Universal Robots URScript: horizontal_swab_path.script

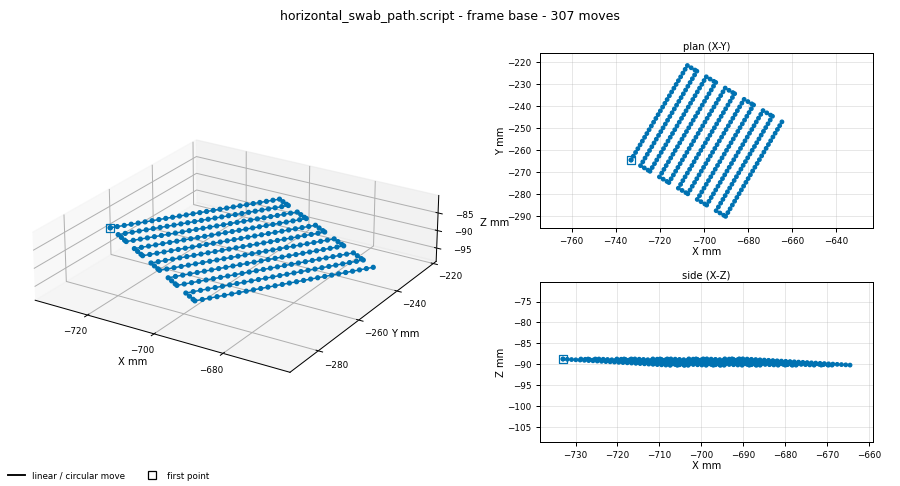
[picture p0: tool path of horizontal_swab_path.script in frame base, 307 of 307 moves have a stored position in this frame; points joined in program order, loops and branches not executed]
def horizontal_swab_path():

  # Move to first swab point perpendicular
  movel(p[-0.73300831, -0.26450111, -0.08872548, -0.83237244, -3.02179964, 0.04578505], a=0.2000, v=0.0300, r=0.0000)

  # Incline tool while keeping TCP XYZ fixed
  movel(p[-0.73300831, -0.26450111, -0.08872548, -0.64311438, -2.27932698, -0.22586576], a=0.1000, v=0.0150, r=0.0000)
  # Horizontal waypoint 1
  movel(p[-0.73198462, -0.26278399, -0.08878548, -0.64311438, -2.27932698, -0.22586576], a=0.1500, v=0.0200, r=0.0000)
  # Horizontal waypoint 2
  movel(p[-0.73096094, -0.26106688, -0.08884547, -0.64311438, -2.27932698, -0.22586576], a=0.1500, v=0.0200, r=0.0000)
  # Horizontal waypoint 3
  movel(p[-0.72993725, -0.25934977, -0.08890546, -0.64311438, -2.27932698, -0.22586576], a=0.1500, v=0.0200, r=0.0000)
  # Horizontal waypoint 4
  movel(p[-0.72891357, -0.25763266, -0.08896545, -0.64311438, -2.27932698, -0.22586576], a=0.1500, v=0.0200, r=0.0000)
  # Horizontal waypoint 5
  movel(p[-0.72788988, -0.25591555, -0.08902544, -0.64311438, -2.27932698, -0.22586576], a=0.1500, v=0.0200, r=0.0000)
  # Horizontal waypoint 6
  movel(p[-0.72686620, -0.25419844, -0.08908543, -0.64311438, -2.27932698, -0.22586576], a=0.1500, v=0.0200, r=0.0000)
  # Horizontal waypoint 7
  movel(p[-0.72584251, -0.25248133, -0.08914542, -0.64311438, -2.27932698, -0.22586576], a=0.1500, v=0.0200, r=0.0000)
  # Horizontal waypoint 8
  movel(p[-0.72481883, -0.25076422, -0.08920541, -0.64311438, -2.27932698, -0.22586576], a=0.1500, v=0.0200, r=0.0000)
  # Horizontal waypoint 9
  movel(p[-0.72379514, -0.24904710, -0.08926540, -0.64311438, -2.27932698, -0.22586576], a=0.1500, v=0.0200, r=0.0000)
  # Horizontal waypoint 10
  movel(p[-0.72277146, -0.24732999, -0.08932539, -0.64311438, -2.27932698, -0.22586576], a=0.1500, v=0.0200, r=0.0000)
  # Horizontal waypoint 11
  movel(p[-0.72174777, -0.24561288, -0.08938538, -0.64311438, -2.27932698, -0.22586576], a=0.1500, v=0.0200, r=0.0000)
  # Horizontal waypoint 12
  movel(p[-0.72072409, -0.24389577, -0.08944538, -0.64311438, -2.27932698, -0.22586576], a=0.1500, v=0.0200, r=0.0000)
  # Horizontal waypoint 13
  movel(p[-0.71970040, -0.24217866, -0.08950537, -0.64311438, -2.27932698, -0.22586576], a=0.1500, v=0.0200, r=0.0000)
  # Horizontal waypoint 14
  movel(p[-0.71867672, -0.24046155, -0.08956536, -0.64311438, -2.27932698, -0.22586576], a=0.1500, v=0.0200, r=0.0000)
  # Horizontal waypoint 15
  movel(p[-0.71765303, -0.23874444, -0.08962535, -0.64311438, -2.27932698, -0.22586576], a=0.1500, v=0.0200, r=0.0000)
  # Horizontal waypoint 16
  movel(p[-0.71662935, -0.23702733, -0.08968534, -0.64311438, -2.27932698, -0.22586576], a=0.1500, v=0.0200, r=0.0000)
  # Horizontal waypoint 17
  movel(p[-0.71560566, -0.23531022, -0.08974533, -0.64311438, -2.27932698, -0.22586576], a=0.1500, v=0.0200, r=0.0000)
  # Horizontal waypoint 18
  movel(p[-0.71458198, -0.23359311, -0.08980532, -0.64311438, -2.27932698, -0.22586576], a=0.1500, v=0.0200, r=0.0000)
  # Horizontal waypoint 19
  movel(p[-0.71355829, -0.23187600, -0.08986531, -0.64311438, -2.27932698, -0.22586576], a=0.1500, v=0.0200, r=0.0000)
  # Horizontal waypoint 20
  movel(p[-0.71253461, -0.23015888, -0.08992530, -0.64311438, -2.27932698, -0.22586576], a=0.1500, v=0.0200, r=0.0000)
  # Horizontal waypoint 21
  movel(p[-0.71151092, -0.22844177, -0.08998530, -0.64311438, -2.27932698, -0.22586576], a=0.1500, v=0.0200, r=0.0000)
  # Horizontal waypoint 22
  movel(p[-0.71048724, -0.22672466, -0.09004529, -0.64311438, -2.27932698, -0.22586576], a=0.1500, v=0.0200, r=0.0000)
  # Horizontal waypoint 23
  movel(p[-0.70946356, -0.22500755, -0.09010528, -0.64311438, -2.27932698, -0.22586576], a=0.1500, v=0.0200, r=0.0000)
  # Horizontal waypoint 24
  movel(p[-0.70843987, -0.22329044, -0.09016527, -0.64311438, -2.27932698, -0.22586576], a=0.1500, v=0.0200, r=0.0000)
  # Horizontal waypoint 25
  movel(p[-0.70741619, -0.22157333, -0.09022526, -0.64311438, -2.27932698, -0.22586576], a=0.1500, v=0.0200, r=0.0000)
  # Horizontal waypoint 26
  movel(p[-0.70569827, -0.22259742, -0.09022307, -0.64311438, -2.27932698, -0.22586576], a=0.1500, v=0.0200, r=0.0000)
  # Horizontal waypoint 27
  movel(p[-0.70398035, -0.22362151, -0.09022089, -0.64311438, -2.27932698, -0.22586576], a=0.1500, v=0.0200, r=0.0000)
  # Horizontal waypoint 28
  movel(p[-0.70312139, -0.22413355, -0.09021980, -0.64311438, -2.27932698, -0.22586576], a=0.1500, v=0.0200, r=0.0000)
  # Horizontal waypoint 29
  movel(p[-0.70414508, -0.22585066, -0.09015981, -0.64311438, -2.27932698, -0.22586576], a=0.1500, v=0.0200, r=0.0000)
  # Horizontal waypoint 30
  movel(p[-0.70516876, -0.22756777, -0.09009982, -0.64311438, -2.27932698, -0.22586576], a=0.1500, v=0.0200, r=0.0000)
  # Horizontal waypoint 31
  movel(p[-0.70619245, -0.22928488, -0.09003983, -0.64311438, -2.27932698, -0.22586576], a=0.1500, v=0.0200, r=0.0000)
  # Horizontal waypoint 32
  movel(p[-0.70721613, -0.23100199, -0.08997983, -0.64311438, -2.27932698, -0.22586576], a=0.1500, v=0.0200, r=0.0000)
  # Horizontal waypoint 33
  movel(p[-0.70823982, -0.23271911, -0.08991984, -0.64311438, -2.27932698, -0.22586576], a=0.1500, v=0.0200, r=0.0000)
  # Horizontal waypoint 34
  movel(p[-0.70926350, -0.23443622, -0.08985985, -0.64311438, -2.27932698, -0.22586576], a=0.1500, v=0.0200, r=0.0000)
  # Horizontal waypoint 35
  movel(p[-0.71028719, -0.23615333, -0.08979986, -0.64311438, -2.27932698, -0.22586576], a=0.1500, v=0.0200, r=0.0000)
  # Horizontal waypoint 36
  movel(p[-0.71131087, -0.23787044, -0.08973987, -0.64311438, -2.27932698, -0.22586576], a=0.1500, v=0.0200, r=0.0000)
  # Horizontal waypoint 37
  movel(p[-0.71233456, -0.23958755, -0.08967988, -0.64311438, -2.27932698, -0.22586576], a=0.1500, v=0.0200, r=0.0000)
  # Horizontal waypoint 38
  movel(p[-0.71335824, -0.24130466, -0.08961989, -0.64311438, -2.27932698, -0.22586576], a=0.1500, v=0.0200, r=0.0000)
  # Horizontal waypoint 39
  movel(p[-0.71438193, -0.24302177, -0.08955990, -0.64311438, -2.27932698, -0.22586576], a=0.1500, v=0.0200, r=0.0000)
  # Horizontal waypoint 40
  movel(p[-0.71540561, -0.24473888, -0.08949991, -0.64311438, -2.27932698, -0.22586576], a=0.1500, v=0.0200, r=0.0000)
  # Horizontal waypoint 41
  movel(p[-0.71642930, -0.24645599, -0.08943991, -0.64311438, -2.27932698, -0.22586576], a=0.1500, v=0.0200, r=0.0000)
  # Horizontal waypoint 42
  movel(p[-0.71745298, -0.24817311, -0.08937992, -0.64311438, -2.27932698, -0.22586576], a=0.1500, v=0.0200, r=0.0000)
  # Horizontal waypoint 43
  movel(p[-0.71847667, -0.24989022, -0.08931993, -0.64311438, -2.27932698, -0.22586576], a=0.1500, v=0.0200, r=0.0000)
  # Horizontal waypoint 44
  movel(p[-0.71950035, -0.25160733, -0.08925994, -0.64311438, -2.27932698, -0.22586576], a=0.1500, v=0.0200, r=0.0000)
  # Horizontal waypoint 45
  movel(p[-0.72052404, -0.25332444, -0.08919995, -0.64311438, -2.27932698, -0.22586576], a=0.1500, v=0.0200, r=0.0000)
  # Horizontal waypoint 46
  movel(p[-0.72154772, -0.25504155, -0.08913996, -0.64311438, -2.27932698, -0.22586576], a=0.1500, v=0.0200, r=0.0000)
  # Horizontal waypoint 47
  movel(p[-0.72257141, -0.25675866, -0.08907997, -0.64311438, -2.27932698, -0.22586576], a=0.1500, v=0.0200, r=0.0000)
  # Horizontal waypoint 48
  movel(p[-0.72359509, -0.25847577, -0.08901998, -0.64311438, -2.27932698, -0.22586576], a=0.1500, v=0.0200, r=0.0000)
  # Horizontal waypoint 49
  movel(p[-0.72461878, -0.26019288, -0.08895999, -0.64311438, -2.27932698, -0.22586576], a=0.1500, v=0.0200, r=0.0000)
  # Horizontal waypoint 50
  movel(p[-0.72564246, -0.26190999, -0.08890000, -0.64311438, -2.27932698, -0.22586576], a=0.1500, v=0.0200, r=0.0000)
  # Horizontal waypoint 51
  movel(p[-0.72666615, -0.26362710, -0.08884000, -0.64311438, -2.27932698, -0.22586576], a=0.1500, v=0.0200, r=0.0000)
  # Horizontal waypoint 52
  movel(p[-0.72768983, -0.26534422, -0.08878001, -0.64311438, -2.27932698, -0.22586576], a=0.1500, v=0.0200, r=0.0000)
  # Horizontal waypoint 53
  movel(p[-0.72871352, -0.26706133, -0.08872002, -0.64311438, -2.27932698, -0.22586576], a=0.1500, v=0.0200, r=0.0000)
  # Horizontal waypoint 54
  movel(p[-0.72699560, -0.26808541, -0.08871784, -0.64311438, -2.27932698, -0.22586576], a=0.1500, v=0.0200, r=0.0000)
  # Horizontal waypoint 55
  movel(p[-0.72527768, -0.26910950, -0.08871566, -0.64311438, -2.27932698, -0.22586576], a=0.1500, v=0.0200, r=0.0000)
  # Horizontal waypoint 56
  movel(p[-0.72441872, -0.26962155, -0.08871456, -0.64311438, -2.27932698, -0.22586576], a=0.1500, v=0.0200, r=0.0000)
  # Horizontal waypoint 57
  movel(p[-0.72339504, -0.26790444, -0.08877455, -0.64311438, -2.27932698, -0.22586576], a=0.1500, v=0.0200, r=0.0000)
  # Horizontal waypoint 58
  movel(p[-0.72237135, -0.26618733, -0.08883455, -0.64311438, -2.27932698, -0.22586576], a=0.1500, v=0.0200, r=0.0000)
  # Horizontal waypoint 59
  movel(p[-0.72134767, -0.26447022, -0.08889454, -0.64311438, -2.27932698, -0.22586576], a=0.1500, v=0.0200, r=0.0000)
  # Horizontal waypoint 60
  movel(p[-0.72032398, -0.26275310, -0.08895453, -0.64311438, -2.27932698, -0.22586576], a=0.1500, v=0.0200, r=0.0000)
  # Horizontal waypoint 61
  movel(p[-0.71930030, -0.26103599, -0.08901452, -0.64311438, -2.27932698, -0.22586576], a=0.1500, v=0.0200, r=0.0000)
  # Horizontal waypoint 62
  movel(p[-0.71827661, -0.25931888, -0.08907451, -0.64311438, -2.27932698, -0.22586576], a=0.1500, v=0.0200, r=0.0000)
  # Horizontal waypoint 63
  movel(p[-0.71725293, -0.25760177, -0.08913450, -0.64311438, -2.27932698, -0.22586576], a=0.1500, v=0.0200, r=0.0000)
  # Horizontal waypoint 64
  movel(p[-0.71622924, -0.25588466, -0.08919449, -0.64311438, -2.27932698, -0.22586576], a=0.1500, v=0.0200, r=0.0000)
  # Horizontal waypoint 65
  movel(p[-0.71520556, -0.25416755, -0.08925448, -0.64311438, -2.27932698, -0.22586576], a=0.1500, v=0.0200, r=0.0000)
  # Horizontal waypoint 66
  movel(p[-0.71418187, -0.25245044, -0.08931447, -0.64311438, -2.27932698, -0.22586576], a=0.1500, v=0.0200, r=0.0000)
  # Horizontal waypoint 67
  movel(p[-0.71315819, -0.25073333, -0.08937446, -0.64311438, -2.27932698, -0.22586576], a=0.1500, v=0.0200, r=0.0000)
  # Horizontal waypoint 68
  movel(p[-0.71213450, -0.24901622, -0.08943445, -0.64311438, -2.27932698, -0.22586576], a=0.1500, v=0.0200, r=0.0000)
  # Horizontal waypoint 69
  movel(p[-0.71111082, -0.24729910, -0.08949445, -0.64311438, -2.27932698, -0.22586576], a=0.1500, v=0.0200, r=0.0000)
  # Horizontal waypoint 70
  movel(p[-0.71008714, -0.24558199, -0.08955444, -0.64311438, -2.27932698, -0.22586576], a=0.1500, v=0.0200, r=0.0000)
  # Horizontal waypoint 71
  movel(p[-0.70906345, -0.24386488, -0.08961443, -0.64311438, -2.27932698, -0.22586576], a=0.1500, v=0.0200, r=0.0000)
  # Horizontal waypoint 72
  movel(p[-0.70803977, -0.24214777, -0.08967442, -0.64311438, -2.27932698, -0.22586576], a=0.1500, v=0.0200, r=0.0000)
  # Horizontal waypoint 73
  movel(p[-0.70701608, -0.24043066, -0.08973441, -0.64311438, -2.27932698, -0.22586576], a=0.1500, v=0.0200, r=0.0000)
  # Horizontal waypoint 74
  movel(p[-0.70599240, -0.23871355, -0.08979440, -0.64311438, -2.27932698, -0.22586576], a=0.1500, v=0.0200, r=0.0000)
  # Horizontal waypoint 75
  movel(p[-0.70496871, -0.23699644, -0.08985439, -0.64311438, -2.27932698, -0.22586576], a=0.1500, v=0.0200, r=0.0000)
  # Horizontal waypoint 76
  movel(p[-0.70394503, -0.23527933, -0.08991438, -0.64311438, -2.27932698, -0.22586576], a=0.1500, v=0.0200, r=0.0000)
  # Horizontal waypoint 77
  movel(p[-0.70292134, -0.23356222, -0.08997437, -0.64311438, -2.27932698, -0.22586576], a=0.1500, v=0.0200, r=0.0000)
  # Horizontal waypoint 78
  movel(p[-0.70189766, -0.23184511, -0.09003437, -0.64311438, -2.27932698, -0.22586576], a=0.1500, v=0.0200, r=0.0000)
  # Horizontal waypoint 79
  movel(p[-0.70087397, -0.23012800, -0.09009436, -0.64311438, -2.27932698, -0.22586576], a=0.1500, v=0.0200, r=0.0000)
  # Horizontal waypoint 80
  movel(p[-0.69985029, -0.22841088, -0.09015435, -0.64311438, -2.27932698, -0.22586576], a=0.1500, v=0.0200, r=0.0000)
  # Horizontal waypoint 81
  movel(p[-0.69882660, -0.22669377, -0.09021434, -0.64311438, -2.27932698, -0.22586576], a=0.1500, v=0.0200, r=0.0000)
  # Horizontal waypoint 82
  movel(p[-0.69710869, -0.22771786, -0.09021215, -0.64311438, -2.27932698, -0.22586576], a=0.1500, v=0.0200, r=0.0000)
  # Horizontal waypoint 83
  movel(p[-0.69539077, -0.22874195, -0.09020997, -0.64311438, -2.27932698, -0.22586576], a=0.1500, v=0.0200, r=0.0000)
  # Horizontal waypoint 84
  movel(p[-0.69453181, -0.22925399, -0.09020888, -0.64311438, -2.27932698, -0.22586576], a=0.1500, v=0.0200, r=0.0000)
  # Horizontal waypoint 85
  movel(p[-0.69555550, -0.23097111, -0.09014889, -0.64311438, -2.27932698, -0.22586576], a=0.1500, v=0.0200, r=0.0000)
  # Horizontal waypoint 86
  movel(p[-0.69657918, -0.23268822, -0.09008890, -0.64311438, -2.27932698, -0.22586576], a=0.1500, v=0.0200, r=0.0000)
  # Horizontal waypoint 87
  movel(p[-0.69760287, -0.23440533, -0.09002890, -0.64311438, -2.27932698, -0.22586576], a=0.1500, v=0.0200, r=0.0000)
  # Horizontal waypoint 88
  movel(p[-0.69862655, -0.23612244, -0.08996891, -0.64311438, -2.27932698, -0.22586576], a=0.1500, v=0.0200, r=0.0000)
  # Horizontal waypoint 89
  movel(p[-0.69965024, -0.23783955, -0.08990892, -0.64311438, -2.27932698, -0.22586576], a=0.1500, v=0.0200, r=0.0000)
  # Horizontal waypoint 90
  movel(p[-0.70067392, -0.23955666, -0.08984893, -0.64311438, -2.27932698, -0.22586576], a=0.1500, v=0.0200, r=0.0000)
  # Horizontal waypoint 91
  movel(p[-0.70169761, -0.24127377, -0.08978894, -0.64311438, -2.27932698, -0.22586576], a=0.1500, v=0.0200, r=0.0000)
  # Horizontal waypoint 92
  movel(p[-0.70272129, -0.24299088, -0.08972895, -0.64311438, -2.27932698, -0.22586576], a=0.1500, v=0.0200, r=0.0000)
  # Horizontal waypoint 93
  movel(p[-0.70374497, -0.24470799, -0.08966896, -0.64311438, -2.27932698, -0.22586576], a=0.1500, v=0.0200, r=0.0000)
  # Horizontal waypoint 94
  movel(p[-0.70476866, -0.24642511, -0.08960897, -0.64311438, -2.27932698, -0.22586576], a=0.1500, v=0.0200, r=0.0000)
  # Horizontal waypoint 95
  movel(p[-0.70579234, -0.24814222, -0.08954898, -0.64311438, -2.27932698, -0.22586576], a=0.1500, v=0.0200, r=0.0000)
  # Horizontal waypoint 96
  movel(p[-0.70681603, -0.24985933, -0.08948898, -0.64311438, -2.27932698, -0.22586576], a=0.1500, v=0.0200, r=0.0000)
  # Horizontal waypoint 97
  movel(p[-0.70783971, -0.25157644, -0.08942899, -0.64311438, -2.27932698, -0.22586576], a=0.1500, v=0.0200, r=0.0000)
  # Horizontal waypoint 98
  movel(p[-0.70886340, -0.25329355, -0.08936900, -0.64311438, -2.27932698, -0.22586576], a=0.1500, v=0.0200, r=0.0000)
  # Horizontal waypoint 99
  movel(p[-0.70988708, -0.25501066, -0.08930901, -0.64311438, -2.27932698, -0.22586576], a=0.1500, v=0.0200, r=0.0000)
  # Horizontal waypoint 100
  movel(p[-0.71091077, -0.25672777, -0.08924902, -0.64311438, -2.27932698, -0.22586576], a=0.1500, v=0.0200, r=0.0000)
  # Horizontal waypoint 101
  movel(p[-0.71193445, -0.25844488, -0.08918903, -0.64311438, -2.27932698, -0.22586576], a=0.1500, v=0.0200, r=0.0000)
  # Horizontal waypoint 102
  movel(p[-0.71295814, -0.26016199, -0.08912904, -0.64311438, -2.27932698, -0.22586576], a=0.1500, v=0.0200, r=0.0000)
  # Horizontal waypoint 103
  movel(p[-0.71398182, -0.26187910, -0.08906905, -0.64311438, -2.27932698, -0.22586576], a=0.1500, v=0.0200, r=0.0000)
  # Horizontal waypoint 104
  movel(p[-0.71500551, -0.26359622, -0.08900906, -0.64311438, -2.27932698, -0.22586576], a=0.1500, v=0.0200, r=0.0000)
  # Horizontal waypoint 105
  movel(p[-0.71602919, -0.26531333, -0.08894907, -0.64311438, -2.27932698, -0.22586576], a=0.1500, v=0.0200, r=0.0000)
  # Horizontal waypoint 106
  movel(p[-0.71705288, -0.26703044, -0.08888907, -0.64311438, -2.27932698, -0.22586576], a=0.1500, v=0.0200, r=0.0000)
  # Horizontal waypoint 107
  movel(p[-0.71807656, -0.26874755, -0.08882908, -0.64311438, -2.27932698, -0.22586576], a=0.1500, v=0.0200, r=0.0000)
  # Horizontal waypoint 108
  movel(p[-0.71910025, -0.27046466, -0.08876909, -0.64311438, -2.27932698, -0.22586576], a=0.1500, v=0.0200, r=0.0000)
  # Horizontal waypoint 109
  movel(p[-0.72012393, -0.27218177, -0.08870910, -0.64311438, -2.27932698, -0.22586576], a=0.1500, v=0.0200, r=0.0000)
  # Horizontal waypoint 110
  movel(p[-0.71840602, -0.27320586, -0.08870692, -0.64311438, -2.27932698, -0.22586576], a=0.1500, v=0.0200, r=0.0000)
  # Horizontal waypoint 111
  movel(p[-0.71668810, -0.27422995, -0.08870473, -0.64311438, -2.27932698, -0.22586576], a=0.1500, v=0.0200, r=0.0000)
  # Horizontal waypoint 112
  movel(p[-0.71582914, -0.27474199, -0.08870364, -0.64311438, -2.27932698, -0.22586576], a=0.1500, v=0.0200, r=0.0000)
  # Horizontal waypoint 113
  movel(p[-0.71480546, -0.27302488, -0.08876363, -0.64311438, -2.27932698, -0.22586576], a=0.1500, v=0.0200, r=0.0000)
  # Horizontal waypoint 114
  movel(p[-0.71378177, -0.27130777, -0.08882362, -0.64311438, -2.27932698, -0.22586576], a=0.1500, v=0.0200, r=0.0000)
  # Horizontal waypoint 115
  movel(p[-0.71275809, -0.26959066, -0.08888361, -0.64311438, -2.27932698, -0.22586576], a=0.1500, v=0.0200, r=0.0000)
  # Horizontal waypoint 116
  movel(p[-0.71173440, -0.26787355, -0.08894360, -0.64311438, -2.27932698, -0.22586576], a=0.1500, v=0.0200, r=0.0000)
  # Horizontal waypoint 117
  movel(p[-0.71071072, -0.26615644, -0.08900360, -0.64311438, -2.27932698, -0.22586576], a=0.1500, v=0.0200, r=0.0000)
  # Horizontal waypoint 118
  movel(p[-0.70968703, -0.26443933, -0.08906359, -0.64311438, -2.27932698, -0.22586576], a=0.1500, v=0.0200, r=0.0000)
  # Horizontal waypoint 119
  movel(p[-0.70866335, -0.26272221, -0.08912358, -0.64311438, -2.27932698, -0.22586576], a=0.1500, v=0.0200, r=0.0000)
  # Horizontal waypoint 120
  movel(p[-0.70763966, -0.26100510, -0.08918357, -0.64311438, -2.27932698, -0.22586576], a=0.1500, v=0.0200, r=0.0000)
  # Horizontal waypoint 121
  movel(p[-0.70661598, -0.25928799, -0.08924356, -0.64311438, -2.27932698, -0.22586576], a=0.1500, v=0.0200, r=0.0000)
  # Horizontal waypoint 122
  movel(p[-0.70559229, -0.25757088, -0.08930355, -0.64311438, -2.27932698, -0.22586576], a=0.1500, v=0.0200, r=0.0000)
  # Horizontal waypoint 123
  movel(p[-0.70456861, -0.25585377, -0.08936354, -0.64311438, -2.27932698, -0.22586576], a=0.1500, v=0.0200, r=0.0000)
  # Horizontal waypoint 124
  movel(p[-0.70354492, -0.25413666, -0.08942353, -0.64311438, -2.27932698, -0.22586576], a=0.1500, v=0.0200, r=0.0000)
  # Horizontal waypoint 125
  movel(p[-0.70252124, -0.25241955, -0.08948352, -0.64311438, -2.27932698, -0.22586576], a=0.1500, v=0.0200, r=0.0000)
  # Horizontal waypoint 126
  movel(p[-0.70149755, -0.25070244, -0.08954352, -0.64311438, -2.27932698, -0.22586576], a=0.1500, v=0.0200, r=0.0000)
  # Horizontal waypoint 127
  movel(p[-0.70047387, -0.24898533, -0.08960351, -0.64311438, -2.27932698, -0.22586576], a=0.1500, v=0.0200, r=0.0000)
  # Horizontal waypoint 128
  movel(p[-0.69945018, -0.24726822, -0.08966350, -0.64311438, -2.27932698, -0.22586576], a=0.1500, v=0.0200, r=0.0000)
  # Horizontal waypoint 129
  movel(p[-0.69842650, -0.24555110, -0.08972349, -0.64311438, -2.27932698, -0.22586576], a=0.1500, v=0.0200, r=0.0000)
  # Horizontal waypoint 130
  movel(p[-0.69740281, -0.24383399, -0.08978348, -0.64311438, -2.27932698, -0.22586576], a=0.1500, v=0.0200, r=0.0000)
  # Horizontal waypoint 131
  movel(p[-0.69637913, -0.24211688, -0.08984347, -0.64311438, -2.27932698, -0.22586576], a=0.1500, v=0.0200, r=0.0000)
  # Horizontal waypoint 132
  movel(p[-0.69535544, -0.24039977, -0.08990346, -0.64311438, -2.27932698, -0.22586576], a=0.1500, v=0.0200, r=0.0000)
  # Horizontal waypoint 133
  movel(p[-0.69433176, -0.23868266, -0.08996345, -0.64311438, -2.27932698, -0.22586576], a=0.1500, v=0.0200, r=0.0000)
  # Horizontal waypoint 134
  movel(p[-0.69330807, -0.23696555, -0.09002344, -0.64311438, -2.27932698, -0.22586576], a=0.1500, v=0.0200, r=0.0000)
  # Horizontal waypoint 135
  movel(p[-0.69228439, -0.23524844, -0.09008343, -0.64311438, -2.27932698, -0.22586576], a=0.1500, v=0.0200, r=0.0000)
  # Horizontal waypoint 136
  movel(p[-0.69126070, -0.23353133, -0.09014342, -0.64311438, -2.27932698, -0.22586576], a=0.1500, v=0.0200, r=0.0000)
  # Horizontal waypoint 137
  movel(p[-0.69023702, -0.23181422, -0.09020342, -0.64311438, -2.27932698, -0.22586576], a=0.1500, v=0.0200, r=0.0000)
  # Horizontal waypoint 138
  movel(p[-0.68851910, -0.23283830, -0.09020123, -0.64311438, -2.27932698, -0.22586576], a=0.1500, v=0.0200, r=0.0000)
  # Horizontal waypoint 139
  movel(p[-0.68680119, -0.23386239, -0.09019905, -0.64311438, -2.27932698, -0.22586576], a=0.1500, v=0.0200, r=0.0000)
  # Horizontal waypoint 140
  movel(p[-0.68594223, -0.23437444, -0.09019795, -0.64311438, -2.27932698, -0.22586576], a=0.1500, v=0.0200, r=0.0000)
  # Horizontal waypoint 141
  movel(p[-0.68696591, -0.23609155, -0.09013796, -0.64311438, -2.27932698, -0.22586576], a=0.1500, v=0.0200, r=0.0000)
  # Horizontal waypoint 142
  movel(p[-0.68798960, -0.23780866, -0.09007797, -0.64311438, -2.27932698, -0.22586576], a=0.1500, v=0.0200, r=0.0000)
  # Horizontal waypoint 143
  movel(p[-0.68901328, -0.23952577, -0.09001798, -0.64311438, -2.27932698, -0.22586576], a=0.1500, v=0.0200, r=0.0000)
  # Horizontal waypoint 144
  movel(p[-0.69003697, -0.24124288, -0.08995799, -0.64311438, -2.27932698, -0.22586576], a=0.1500, v=0.0200, r=0.0000)
  # Horizontal waypoint 145
  movel(p[-0.69106065, -0.24295999, -0.08989800, -0.64311438, -2.27932698, -0.22586576], a=0.1500, v=0.0200, r=0.0000)
  # Horizontal waypoint 146
  movel(p[-0.69208434, -0.24467711, -0.08983801, -0.64311438, -2.27932698, -0.22586576], a=0.1500, v=0.0200, r=0.0000)
  # Horizontal waypoint 147
  movel(p[-0.69310802, -0.24639422, -0.08977802, -0.64311438, -2.27932698, -0.22586576], a=0.1500, v=0.0200, r=0.0000)
  # Horizontal waypoint 148
  movel(p[-0.69413171, -0.24811133, -0.08971803, -0.64311438, -2.27932698, -0.22586576], a=0.1500, v=0.0200, r=0.0000)
  # Horizontal waypoint 149
  movel(p[-0.69515539, -0.24982844, -0.08965804, -0.64311438, -2.27932698, -0.22586576], a=0.1500, v=0.0200, r=0.0000)
  # Horizontal waypoint 150
  movel(p[-0.69617908, -0.25154555, -0.08959805, -0.64311438, -2.27932698, -0.22586576], a=0.1500, v=0.0200, r=0.0000)
  # Horizontal waypoint 151
  movel(p[-0.69720276, -0.25326266, -0.08953805, -0.64311438, -2.27932698, -0.22586576], a=0.1500, v=0.0200, r=0.0000)
  # Horizontal waypoint 152
  movel(p[-0.69822645, -0.25497977, -0.08947806, -0.64311438, -2.27932698, -0.22586576], a=0.1500, v=0.0200, r=0.0000)
  # Horizontal waypoint 153
  movel(p[-0.69925013, -0.25669688, -0.08941807, -0.64311438, -2.27932698, -0.22586576], a=0.1500, v=0.0200, r=0.0000)
  # Horizontal waypoint 154
  movel(p[-0.70027382, -0.25841399, -0.08935808, -0.64311438, -2.27932698, -0.22586576], a=0.1500, v=0.0200, r=0.0000)
  # Horizontal waypoint 155
  movel(p[-0.70129750, -0.26013110, -0.08929809, -0.64311438, -2.27932698, -0.22586576], a=0.1500, v=0.0200, r=0.0000)
  # Horizontal waypoint 156
  movel(p[-0.70232119, -0.26184821, -0.08923810, -0.64311438, -2.27932698, -0.22586576], a=0.1500, v=0.0200, r=0.0000)
  # Horizontal waypoint 157
  movel(p[-0.70334487, -0.26356533, -0.08917811, -0.64311438, -2.27932698, -0.22586576], a=0.1500, v=0.0200, r=0.0000)
  # Horizontal waypoint 158
  movel(p[-0.70436855, -0.26528244, -0.08911812, -0.64311438, -2.27932698, -0.22586576], a=0.1500, v=0.0200, r=0.0000)
  # Horizontal waypoint 159
  movel(p[-0.70539224, -0.26699955, -0.08905813, -0.64311438, -2.27932698, -0.22586576], a=0.1500, v=0.0200, r=0.0000)
  # Horizontal waypoint 160
  movel(p[-0.70641592, -0.26871666, -0.08899814, -0.64311438, -2.27932698, -0.22586576], a=0.1500, v=0.0200, r=0.0000)
  # Horizontal waypoint 161
  movel(p[-0.70743961, -0.27043377, -0.08893814, -0.64311438, -2.27932698, -0.22586576], a=0.1500, v=0.0200, r=0.0000)
  # Horizontal waypoint 162
  movel(p[-0.70846330, -0.27215088, -0.08887815, -0.64311438, -2.27932698, -0.22586576], a=0.1500, v=0.0200, r=0.0000)
  # Horizontal waypoint 163
  movel(p[-0.70948698, -0.27386799, -0.08881816, -0.64311438, -2.27932698, -0.22586576], a=0.1500, v=0.0200, r=0.0000)
  # Horizontal waypoint 164
  movel(p[-0.71051067, -0.27558510, -0.08875817, -0.64311438, -2.27932698, -0.22586576], a=0.1500, v=0.0200, r=0.0000)
  # Horizontal waypoint 165
  movel(p[-0.71153435, -0.27730222, -0.08869818, -0.64311438, -2.27932698, -0.22586576], a=0.1500, v=0.0200, r=0.0000)
  # Horizontal waypoint 166
  movel(p[-0.70981643, -0.27832630, -0.08869600, -0.64311438, -2.27932698, -0.22586576], a=0.1500, v=0.0200, r=0.0000)
  # Horizontal waypoint 167
  movel(p[-0.70809852, -0.27935039, -0.08869381, -0.64311438, -2.27932698, -0.22586576], a=0.1500, v=0.0200, r=0.0000)
  # Horizontal waypoint 168
  movel(p[-0.70723956, -0.27986244, -0.08869272, -0.64311438, -2.27932698, -0.22586576], a=0.1500, v=0.0200, r=0.0000)
  # Horizontal waypoint 169
  movel(p[-0.70621587, -0.27814533, -0.08875271, -0.64311438, -2.27932698, -0.22586576], a=0.1500, v=0.0200, r=0.0000)
  # Horizontal waypoint 170
  movel(p[-0.70519219, -0.27642821, -0.08881270, -0.64311438, -2.27932698, -0.22586576], a=0.1500, v=0.0200, r=0.0000)
  # Horizontal waypoint 171
  movel(p[-0.70416850, -0.27471110, -0.08887269, -0.64311438, -2.27932698, -0.22586576], a=0.1500, v=0.0200, r=0.0000)
  # Horizontal waypoint 172
  movel(p[-0.70314482, -0.27299399, -0.08893268, -0.64311438, -2.27932698, -0.22586576], a=0.1500, v=0.0200, r=0.0000)
  # Horizontal waypoint 173
  movel(p[-0.70212113, -0.27127688, -0.08899267, -0.64311438, -2.27932698, -0.22586576], a=0.1500, v=0.0200, r=0.0000)
  # Horizontal waypoint 174
  movel(p[-0.70109745, -0.26955977, -0.08905267, -0.64311438, -2.27932698, -0.22586576], a=0.1500, v=0.0200, r=0.0000)
  # Horizontal waypoint 175
  movel(p[-0.70007376, -0.26784266, -0.08911266, -0.64311438, -2.27932698, -0.22586576], a=0.1500, v=0.0200, r=0.0000)
  # Horizontal waypoint 176
  movel(p[-0.69905008, -0.26612555, -0.08917265, -0.64311438, -2.27932698, -0.22586576], a=0.1500, v=0.0200, r=0.0000)
  # Horizontal waypoint 177
  movel(p[-0.69802639, -0.26440844, -0.08923264, -0.64311438, -2.27932698, -0.22586576], a=0.1500, v=0.0200, r=0.0000)
  # Horizontal waypoint 178
  movel(p[-0.69700271, -0.26269133, -0.08929263, -0.64311438, -2.27932698, -0.22586576], a=0.1500, v=0.0200, r=0.0000)
  # Horizontal waypoint 179
  movel(p[-0.69597902, -0.26097422, -0.08935262, -0.64311438, -2.27932698, -0.22586576], a=0.1500, v=0.0200, r=0.0000)
  # Horizontal waypoint 180
  movel(p[-0.69495534, -0.25925710, -0.08941261, -0.64311438, -2.27932698, -0.22586576], a=0.1500, v=0.0200, r=0.0000)
  # Horizontal waypoint 181
  movel(p[-0.69393165, -0.25753999, -0.08947260, -0.64311438, -2.27932698, -0.22586576], a=0.1500, v=0.0200, r=0.0000)
  # Horizontal waypoint 182
  movel(p[-0.69290797, -0.25582288, -0.08953259, -0.64311438, -2.27932698, -0.22586576], a=0.1500, v=0.0200, r=0.0000)
  # Horizontal waypoint 183
  movel(p[-0.69188428, -0.25410577, -0.08959258, -0.64311438, -2.27932698, -0.22586576], a=0.1500, v=0.0200, r=0.0000)
  # Horizontal waypoint 184
  movel(p[-0.69086060, -0.25238866, -0.08965257, -0.64311438, -2.27932698, -0.22586576], a=0.1500, v=0.0200, r=0.0000)
  # Horizontal waypoint 185
  movel(p[-0.68983691, -0.25067155, -0.08971257, -0.64311438, -2.27932698, -0.22586576], a=0.1500, v=0.0200, r=0.0000)
  # Horizontal waypoint 186
  movel(p[-0.68881323, -0.24895444, -0.08977256, -0.64311438, -2.27932698, -0.22586576], a=0.1500, v=0.0200, r=0.0000)
  # Horizontal waypoint 187
  movel(p[-0.68778955, -0.24723733, -0.08983255, -0.64311438, -2.27932698, -0.22586576], a=0.1500, v=0.0200, r=0.0000)
  # Horizontal waypoint 188
  movel(p[-0.68676586, -0.24552022, -0.08989254, -0.64311438, -2.27932698, -0.22586576], a=0.1500, v=0.0200, r=0.0000)
  # Horizontal waypoint 189
  movel(p[-0.68574218, -0.24380310, -0.08995253, -0.64311438, -2.27932698, -0.22586576], a=0.1500, v=0.0200, r=0.0000)
  # Horizontal waypoint 190
  movel(p[-0.68471849, -0.24208599, -0.09001252, -0.64311438, -2.27932698, -0.22586576], a=0.1500, v=0.0200, r=0.0000)
  # Horizontal waypoint 191
  movel(p[-0.68369481, -0.24036888, -0.09007251, -0.64311438, -2.27932698, -0.22586576], a=0.1500, v=0.0200, r=0.0000)
  # Horizontal waypoint 192
  movel(p[-0.68267112, -0.23865177, -0.09013250, -0.64311438, -2.27932698, -0.22586576], a=0.1500, v=0.0200, r=0.0000)
  # Horizontal waypoint 193
  movel(p[-0.68164744, -0.23693466, -0.09019249, -0.64311438, -2.27932698, -0.22586576], a=0.1500, v=0.0200, r=0.0000)
  # Horizontal waypoint 194
  movel(p[-0.67992952, -0.23795875, -0.09019031, -0.64311438, -2.27932698, -0.22586576], a=0.1500, v=0.0200, r=0.0000)
  # Horizontal waypoint 195
  movel(p[-0.67821160, -0.23898284, -0.09018813, -0.64311438, -2.27932698, -0.22586576], a=0.1500, v=0.0200, r=0.0000)
  # Horizontal waypoint 196
  movel(p[-0.67735265, -0.23949488, -0.09018703, -0.64311438, -2.27932698, -0.22586576], a=0.1500, v=0.0200, r=0.0000)
  # Horizontal waypoint 197
  movel(p[-0.67837633, -0.24121199, -0.09012704, -0.64311438, -2.27932698, -0.22586576], a=0.1500, v=0.0200, r=0.0000)
  # Horizontal waypoint 198
  movel(p[-0.67940001, -0.24292911, -0.09006705, -0.64311438, -2.27932698, -0.22586576], a=0.1500, v=0.0200, r=0.0000)
  # Horizontal waypoint 199
  movel(p[-0.68042370, -0.24464622, -0.09000706, -0.64311438, -2.27932698, -0.22586576], a=0.1500, v=0.0200, r=0.0000)
  # Horizontal waypoint 200
  movel(p[-0.68144738, -0.24636333, -0.08994707, -0.64311438, -2.27932698, -0.22586576], a=0.1500, v=0.0200, r=0.0000)
  # Horizontal waypoint 201
  movel(p[-0.68247107, -0.24808044, -0.08988708, -0.64311438, -2.27932698, -0.22586576], a=0.1500, v=0.0200, r=0.0000)
  # Horizontal waypoint 202
  movel(p[-0.68349475, -0.24979755, -0.08982709, -0.64311438, -2.27932698, -0.22586576], a=0.1500, v=0.0200, r=0.0000)
  # Horizontal waypoint 203
  movel(p[-0.68451844, -0.25151466, -0.08976710, -0.64311438, -2.27932698, -0.22586576], a=0.1500, v=0.0200, r=0.0000)
  # Horizontal waypoint 204
  movel(p[-0.68554212, -0.25323177, -0.08970711, -0.64311438, -2.27932698, -0.22586576], a=0.1500, v=0.0200, r=0.0000)
  # Horizontal waypoint 205
  movel(p[-0.68656581, -0.25494888, -0.08964711, -0.64311438, -2.27932698, -0.22586576], a=0.1500, v=0.0200, r=0.0000)
  # Horizontal waypoint 206
  movel(p[-0.68758949, -0.25666599, -0.08958712, -0.64311438, -2.27932698, -0.22586576], a=0.1500, v=0.0200, r=0.0000)
  # Horizontal waypoint 207
  movel(p[-0.68861318, -0.25838310, -0.08952713, -0.64311438, -2.27932698, -0.22586576], a=0.1500, v=0.0200, r=0.0000)
  # Horizontal waypoint 208
  movel(p[-0.68963686, -0.26010022, -0.08946714, -0.64311438, -2.27932698, -0.22586576], a=0.1500, v=0.0200, r=0.0000)
  # Horizontal waypoint 209
  movel(p[-0.69066055, -0.26181733, -0.08940715, -0.64311438, -2.27932698, -0.22586576], a=0.1500, v=0.0200, r=0.0000)
  # Horizontal waypoint 210
  movel(p[-0.69168423, -0.26353444, -0.08934716, -0.64311438, -2.27932698, -0.22586576], a=0.1500, v=0.0200, r=0.0000)
  # Horizontal waypoint 211
  movel(p[-0.69270792, -0.26525155, -0.08928717, -0.64311438, -2.27932698, -0.22586576], a=0.1500, v=0.0200, r=0.0000)
  # Horizontal waypoint 212
  movel(p[-0.69373160, -0.26696866, -0.08922718, -0.64311438, -2.27932698, -0.22586576], a=0.1500, v=0.0200, r=0.0000)
  # Horizontal waypoint 213
  movel(p[-0.69475529, -0.26868577, -0.08916719, -0.64311438, -2.27932698, -0.22586576], a=0.1500, v=0.0200, r=0.0000)
  # Horizontal waypoint 214
  movel(p[-0.69577897, -0.27040288, -0.08910720, -0.64311438, -2.27932698, -0.22586576], a=0.1500, v=0.0200, r=0.0000)
  # Horizontal waypoint 215
  movel(p[-0.69680266, -0.27211999, -0.08904721, -0.64311438, -2.27932698, -0.22586576], a=0.1500, v=0.0200, r=0.0000)
  # Horizontal waypoint 216
  movel(p[-0.69782634, -0.27383710, -0.08898721, -0.64311438, -2.27932698, -0.22586576], a=0.1500, v=0.0200, r=0.0000)
  # Horizontal waypoint 217
  movel(p[-0.69885003, -0.27555421, -0.08892722, -0.64311438, -2.27932698, -0.22586576], a=0.1500, v=0.0200, r=0.0000)
  # Horizontal waypoint 218
  movel(p[-0.69987371, -0.27727133, -0.08886723, -0.64311438, -2.27932698, -0.22586576], a=0.1500, v=0.0200, r=0.0000)
  # Horizontal waypoint 219
  movel(p[-0.70089740, -0.27898844, -0.08880724, -0.64311438, -2.27932698, -0.22586576], a=0.1500, v=0.0200, r=0.0000)
  # Horizontal waypoint 220
  movel(p[-0.70192108, -0.28070555, -0.08874725, -0.64311438, -2.27932698, -0.22586576], a=0.1500, v=0.0200, r=0.0000)
  # Horizontal waypoint 221
  movel(p[-0.70294477, -0.28242266, -0.08868726, -0.64311438, -2.27932698, -0.22586576], a=0.1500, v=0.0200, r=0.0000)
  # Horizontal waypoint 222
  movel(p[-0.70122685, -0.28344675, -0.08868507, -0.64311438, -2.27932698, -0.22586576], a=0.1500, v=0.0200, r=0.0000)
  # Horizontal waypoint 223
  movel(p[-0.69950893, -0.28447084, -0.08868289, -0.64311438, -2.27932698, -0.22586576], a=0.1500, v=0.0200, r=0.0000)
  # Horizontal waypoint 224
  movel(p[-0.69864998, -0.28498288, -0.08868180, -0.64311438, -2.27932698, -0.22586576], a=0.1500, v=0.0200, r=0.0000)
  # Horizontal waypoint 225
  movel(p[-0.69762629, -0.28326577, -0.08874179, -0.64311438, -2.27932698, -0.22586576], a=0.1500, v=0.0200, r=0.0000)
  # Horizontal waypoint 226
  movel(p[-0.69660261, -0.28154866, -0.08880178, -0.64311438, -2.27932698, -0.22586576], a=0.1500, v=0.0200, r=0.0000)
  # Horizontal waypoint 227
  movel(p[-0.69557892, -0.27983155, -0.08886177, -0.64311438, -2.27932698, -0.22586576], a=0.1500, v=0.0200, r=0.0000)
  # Horizontal waypoint 228
  movel(p[-0.69455524, -0.27811444, -0.08892176, -0.64311438, -2.27932698, -0.22586576], a=0.1500, v=0.0200, r=0.0000)
  # Horizontal waypoint 229
  movel(p[-0.69353155, -0.27639733, -0.08898175, -0.64311438, -2.27932698, -0.22586576], a=0.1500, v=0.0200, r=0.0000)
  # Horizontal waypoint 230
  movel(p[-0.69250787, -0.27468021, -0.08904174, -0.64311438, -2.27932698, -0.22586576], a=0.1500, v=0.0200, r=0.0000)
  # Horizontal waypoint 231
  movel(p[-0.69148418, -0.27296310, -0.08910174, -0.64311438, -2.27932698, -0.22586576], a=0.1500, v=0.0200, r=0.0000)
  # Horizontal waypoint 232
  movel(p[-0.69046050, -0.27124599, -0.08916173, -0.64311438, -2.27932698, -0.22586576], a=0.1500, v=0.0200, r=0.0000)
  # Horizontal waypoint 233
  movel(p[-0.68943681, -0.26952888, -0.08922172, -0.64311438, -2.27932698, -0.22586576], a=0.1500, v=0.0200, r=0.0000)
  # Horizontal waypoint 234
  movel(p[-0.68841313, -0.26781177, -0.08928171, -0.64311438, -2.27932698, -0.22586576], a=0.1500, v=0.0200, r=0.0000)
  # Horizontal waypoint 235
  movel(p[-0.68738944, -0.26609466, -0.08934170, -0.64311438, -2.27932698, -0.22586576], a=0.1500, v=0.0200, r=0.0000)
  # Horizontal waypoint 236
  movel(p[-0.68636576, -0.26437755, -0.08940169, -0.64311438, -2.27932698, -0.22586576], a=0.1500, v=0.0200, r=0.0000)
  # Horizontal waypoint 237
  movel(p[-0.68534207, -0.26266044, -0.08946168, -0.64311438, -2.27932698, -0.22586576], a=0.1500, v=0.0200, r=0.0000)
  # Horizontal waypoint 238
  movel(p[-0.68431839, -0.26094333, -0.08952167, -0.64311438, -2.27932698, -0.22586576], a=0.1500, v=0.0200, r=0.0000)
  # Horizontal waypoint 239
  movel(p[-0.68329470, -0.25922621, -0.08958166, -0.64311438, -2.27932698, -0.22586576], a=0.1500, v=0.0200, r=0.0000)
  # Horizontal waypoint 240
  movel(p[-0.68227102, -0.25750910, -0.08964165, -0.64311438, -2.27932698, -0.22586576], a=0.1500, v=0.0200, r=0.0000)
  # Horizontal waypoint 241
  movel(p[-0.68124733, -0.25579199, -0.08970164, -0.64311438, -2.27932698, -0.22586576], a=0.1500, v=0.0200, r=0.0000)
  # Horizontal waypoint 242
  movel(p[-0.68022365, -0.25407488, -0.08976164, -0.64311438, -2.27932698, -0.22586576], a=0.1500, v=0.0200, r=0.0000)
  # Horizontal waypoint 243
  movel(p[-0.67919996, -0.25235777, -0.08982163, -0.64311438, -2.27932698, -0.22586576], a=0.1500, v=0.0200, r=0.0000)
  # Horizontal waypoint 244
  movel(p[-0.67817628, -0.25064066, -0.08988162, -0.64311438, -2.27932698, -0.22586576], a=0.1500, v=0.0200, r=0.0000)
  # Horizontal waypoint 245
  movel(p[-0.67715259, -0.24892355, -0.08994161, -0.64311438, -2.27932698, -0.22586576], a=0.1500, v=0.0200, r=0.0000)
  # Horizontal waypoint 246
  movel(p[-0.67612891, -0.24720644, -0.09000160, -0.64311438, -2.27932698, -0.22586576], a=0.1500, v=0.0200, r=0.0000)
  # Horizontal waypoint 247
  movel(p[-0.67510522, -0.24548933, -0.09006159, -0.64311438, -2.27932698, -0.22586576], a=0.1500, v=0.0200, r=0.0000)
  # Horizontal waypoint 248
  movel(p[-0.67408154, -0.24377222, -0.09012158, -0.64311438, -2.27932698, -0.22586576], a=0.1500, v=0.0200, r=0.0000)
  # Horizontal waypoint 249
  movel(p[-0.67305785, -0.24205510, -0.09018157, -0.64311438, -2.27932698, -0.22586576], a=0.1500, v=0.0200, r=0.0000)
  # Horizontal waypoint 250
  movel(p[-0.67133994, -0.24307919, -0.09017939, -0.64311438, -2.27932698, -0.22586576], a=0.1500, v=0.0200, r=0.0000)
  # Horizontal waypoint 251
  movel(p[-0.66962202, -0.24410328, -0.09017720, -0.64311438, -2.27932698, -0.22586576], a=0.1500, v=0.0200, r=0.0000)
  # Horizontal waypoint 252
  movel(p[-0.66876306, -0.24461533, -0.09017611, -0.64311438, -2.27932698, -0.22586576], a=0.1500, v=0.0200, r=0.0000)
  # Horizontal waypoint 253
  movel(p[-0.66978675, -0.24633244, -0.09011612, -0.64311438, -2.27932698, -0.22586576], a=0.1500, v=0.0200, r=0.0000)
  # Horizontal waypoint 254
  movel(p[-0.67081043, -0.24804955, -0.09005613, -0.64311438, -2.27932698, -0.22586576], a=0.1500, v=0.0200, r=0.0000)
  # Horizontal waypoint 255
  movel(p[-0.67183412, -0.24976666, -0.08999614, -0.64311438, -2.27932698, -0.22586576], a=0.1500, v=0.0200, r=0.0000)
  # Horizontal waypoint 256
  movel(p[-0.67285780, -0.25148377, -0.08993615, -0.64311438, -2.27932698, -0.22586576], a=0.1500, v=0.0200, r=0.0000)
  # Horizontal waypoint 257
  movel(p[-0.67388149, -0.25320088, -0.08987616, -0.64311438, -2.27932698, -0.22586576], a=0.1500, v=0.0200, r=0.0000)
  # Horizontal waypoint 258
  movel(p[-0.67490517, -0.25491799, -0.08981617, -0.64311438, -2.27932698, -0.22586576], a=0.1500, v=0.0200, r=0.0000)
  # Horizontal waypoint 259
  movel(p[-0.67592886, -0.25663510, -0.08975617, -0.64311438, -2.27932698, -0.22586576], a=0.1500, v=0.0200, r=0.0000)
  # Horizontal waypoint 260
  movel(p[-0.67695254, -0.25835221, -0.08969618, -0.64311438, -2.27932698, -0.22586576], a=0.1500, v=0.0200, r=0.0000)
  # Horizontal waypoint 261
  movel(p[-0.67797623, -0.26006933, -0.08963619, -0.64311438, -2.27932698, -0.22586576], a=0.1500, v=0.0200, r=0.0000)
  # Horizontal waypoint 262
  movel(p[-0.67899991, -0.26178644, -0.08957620, -0.64311438, -2.27932698, -0.22586576], a=0.1500, v=0.0200, r=0.0000)
  # Horizontal waypoint 263
  movel(p[-0.68002360, -0.26350355, -0.08951621, -0.64311438, -2.27932698, -0.22586576], a=0.1500, v=0.0200, r=0.0000)
  # Horizontal waypoint 264
  movel(p[-0.68104728, -0.26522066, -0.08945622, -0.64311438, -2.27932698, -0.22586576], a=0.1500, v=0.0200, r=0.0000)
  # Horizontal waypoint 265
  movel(p[-0.68207096, -0.26693777, -0.08939623, -0.64311438, -2.27932698, -0.22586576], a=0.1500, v=0.0200, r=0.0000)
  # Horizontal waypoint 266
  movel(p[-0.68309465, -0.26865488, -0.08933624, -0.64311438, -2.27932698, -0.22586576], a=0.1500, v=0.0200, r=0.0000)
  # Horizontal waypoint 267
  movel(p[-0.68411833, -0.27037199, -0.08927625, -0.64311438, -2.27932698, -0.22586576], a=0.1500, v=0.0200, r=0.0000)
  # Horizontal waypoint 268
  movel(p[-0.68514202, -0.27208910, -0.08921626, -0.64311438, -2.27932698, -0.22586576], a=0.1500, v=0.0200, r=0.0000)
  # Horizontal waypoint 269
  movel(p[-0.68616570, -0.27380621, -0.08915626, -0.64311438, -2.27932698, -0.22586576], a=0.1500, v=0.0200, r=0.0000)
  # Horizontal waypoint 270
  movel(p[-0.68718939, -0.27552332, -0.08909627, -0.64311438, -2.27932698, -0.22586576], a=0.1500, v=0.0200, r=0.0000)
  # Horizontal waypoint 271
  movel(p[-0.68821307, -0.27724044, -0.08903628, -0.64311438, -2.27932698, -0.22586576], a=0.1500, v=0.0200, r=0.0000)
  # Horizontal waypoint 272
  movel(p[-0.68923676, -0.27895755, -0.08897629, -0.64311438, -2.27932698, -0.22586576], a=0.1500, v=0.0200, r=0.0000)
  # Horizontal waypoint 273
  movel(p[-0.69026044, -0.28067466, -0.08891630, -0.64311438, -2.27932698, -0.22586576], a=0.1500, v=0.0200, r=0.0000)
  # Horizontal waypoint 274
  movel(p[-0.69128413, -0.28239177, -0.08885631, -0.64311438, -2.27932698, -0.22586576], a=0.1500, v=0.0200, r=0.0000)
  # Horizontal waypoint 275
  movel(p[-0.69230781, -0.28410888, -0.08879632, -0.64311438, -2.27932698, -0.22586576], a=0.1500, v=0.0200, r=0.0000)
  # Horizontal waypoint 276
  movel(p[-0.69333150, -0.28582599, -0.08873633, -0.64311438, -2.27932698, -0.22586576], a=0.1500, v=0.0200, r=0.0000)
  # Horizontal waypoint 277
  movel(p[-0.69435518, -0.28754310, -0.08867634, -0.64311438, -2.27932698, -0.22586576], a=0.1500, v=0.0200, r=0.0000)
  # Horizontal waypoint 278
  movel(p[-0.69263727, -0.28856719, -0.08867415, -0.64311438, -2.27932698, -0.22586576], a=0.1500, v=0.0200, r=0.0000)
  # Horizontal waypoint 279
  movel(p[-0.69091935, -0.28959128, -0.08867197, -0.64311438, -2.27932698, -0.22586576], a=0.1500, v=0.0200, r=0.0000)
  # Horizontal waypoint 280
  movel(p[-0.69006039, -0.29010333, -0.08867088, -0.64311438, -2.27932698, -0.22586576], a=0.1500, v=0.0200, r=0.0000)
  # Horizontal waypoint 281
  movel(p[-0.68903671, -0.28838621, -0.08873087, -0.64311438, -2.27932698, -0.22586576], a=0.1500, v=0.0200, r=0.0000)
  # Horizontal waypoint 282
  movel(p[-0.68801302, -0.28666910, -0.08879086, -0.64311438, -2.27932698, -0.22586576], a=0.1500, v=0.0200, r=0.0000)
  # Horizontal waypoint 283
  movel(p[-0.68698934, -0.28495199, -0.08885085, -0.64311438, -2.27932698, -0.22586576], a=0.1500, v=0.0200, r=0.0000)
  # Horizontal waypoint 284
  movel(p[-0.68596565, -0.28323488, -0.08891084, -0.64311438, -2.27932698, -0.22586576], a=0.1500, v=0.0200, r=0.0000)
  # Horizontal waypoint 285
  movel(p[-0.68494197, -0.28151777, -0.08897083, -0.64311438, -2.27932698, -0.22586576], a=0.1500, v=0.0200, r=0.0000)
  # Horizontal waypoint 286
  movel(p[-0.68391828, -0.27980066, -0.08903082, -0.64311438, -2.27932698, -0.22586576], a=0.1500, v=0.0200, r=0.0000)
  # Horizontal waypoint 287
  movel(p[-0.68289460, -0.27808355, -0.08909081, -0.64311438, -2.27932698, -0.22586576], a=0.1500, v=0.0200, r=0.0000)
  # Horizontal waypoint 288
  movel(p[-0.68187091, -0.27636644, -0.08915080, -0.64311438, -2.27932698, -0.22586576], a=0.1500, v=0.0200, r=0.0000)
  # Horizontal waypoint 289
  movel(p[-0.68084723, -0.27464932, -0.08921079, -0.64311438, -2.27932698, -0.22586576], a=0.1500, v=0.0200, r=0.0000)
  # Horizontal waypoint 290
  movel(p[-0.67982354, -0.27293221, -0.08927079, -0.64311438, -2.27932698, -0.22586576], a=0.1500, v=0.0200, r=0.0000)
  # Horizontal waypoint 291
  movel(p[-0.67879986, -0.27121510, -0.08933078, -0.64311438, -2.27932698, -0.22586576], a=0.1500, v=0.0200, r=0.0000)
  # Horizontal waypoint 292
  movel(p[-0.67777617, -0.26949799, -0.08939077, -0.64311438, -2.27932698, -0.22586576], a=0.1500, v=0.0200, r=0.0000)
  # Horizontal waypoint 293
  movel(p[-0.67675249, -0.26778088, -0.08945076, -0.64311438, -2.27932698, -0.22586576], a=0.1500, v=0.0200, r=0.0000)
  # Horizontal waypoint 294
  movel(p[-0.67572880, -0.26606377, -0.08951075, -0.64311438, -2.27932698, -0.22586576], a=0.1500, v=0.0200, r=0.0000)
  # Horizontal waypoint 295
  movel(p[-0.67470512, -0.26434666, -0.08957074, -0.64311438, -2.27932698, -0.22586576], a=0.1500, v=0.0200, r=0.0000)
  # Horizontal waypoint 296
  movel(p[-0.67368143, -0.26262955, -0.08963073, -0.64311438, -2.27932698, -0.22586576], a=0.1500, v=0.0200, r=0.0000)
  # Horizontal waypoint 297
  movel(p[-0.67265775, -0.26091244, -0.08969072, -0.64311438, -2.27932698, -0.22586576], a=0.1500, v=0.0200, r=0.0000)
  # Horizontal waypoint 298
  movel(p[-0.67163407, -0.25919533, -0.08975071, -0.64311438, -2.27932698, -0.22586576], a=0.1500, v=0.0200, r=0.0000)
  # Horizontal waypoint 299
  movel(p[-0.67061038, -0.25747822, -0.08981071, -0.64311438, -2.27932698, -0.22586576], a=0.1500, v=0.0200, r=0.0000)
  # Horizontal waypoint 300
  movel(p[-0.66958670, -0.25576110, -0.08987070, -0.64311438, -2.27932698, -0.22586576], a=0.1500, v=0.0200, r=0.0000)
  # Horizontal waypoint 301
  movel(p[-0.66856301, -0.25404399, -0.08993069, -0.64311438, -2.27932698, -0.22586576], a=0.1500, v=0.0200, r=0.0000)
  # Horizontal waypoint 302
  movel(p[-0.66753933, -0.25232688, -0.08999068, -0.64311438, -2.27932698, -0.22586576], a=0.1500, v=0.0200, r=0.0000)
  # Horizontal waypoint 303
  movel(p[-0.66651564, -0.25060977, -0.09005067, -0.64311438, -2.27932698, -0.22586576], a=0.1500, v=0.0200, r=0.0000)
  # Horizontal waypoint 304
  movel(p[-0.66549196, -0.24889266, -0.09011066, -0.64311438, -2.27932698, -0.22586576], a=0.1500, v=0.0200, r=0.0000)
  # Horizontal waypoint 305
  movel(p[-0.66446827, -0.24717555, -0.09017065, -0.64311438, -2.27932698, -0.22586576], a=0.1500, v=0.0200, r=0.0000)
end
